(* IEC 61131-3 sources: rusty/tests/lit/single/polymorphism/fnptr, 14 files *)

(* ---- function_block_call_explicit_arguments.st ---- *)
// RUN: %COMPILE %s && %RUN | %CHECK %s

TYPE Position2D:
    STRUCT
        x: DINT;
        y: DINT;
    END_STRUCT
END_TYPE

FUNCTION_BLOCK FbA
    VAR
        localState: DINT := 0;
    END_VAR

    VAR_INPUT
        in1: DINT;
        in2: STRING;
        in3: Position2D;
        in4: ARRAY[1..2] OF STRING;
        in5: ARRAY[1..2] OF Position2D;
    END_VAR

    VAR_OUTPUT
        out1: DINT;
        out2: STRING;
        out3: Position2D;
        out4: ARRAY[1..2] OF STRING;
        out5: ARRAY[1..2] OF Position2D;
    END_VAR

    VAR_IN_OUT
        inout1: DINT;
        inout2: STRING;
        inout3: Position2D;
        inout4: ARRAY[1..2] OF STRING;
        inout5: ARRAY[1..2] OF Position2D;
    END_VAR

    METHOD increaseLocalState
        localState := localState + 1;
    END_METHOD

    printf('localState = %d$N', localState);

    printf('in1 = %d$N', in1);
    printf('in2 = %s$N', ADR(in2));
    printf('in3 = (%d, %d)$N', in3.x, in3.y);
    printf('in4 = [%s, %s]$N', ADR(in4[1]), ADR(in4[2]));
    printf('in5 = [(%d, %d), (%d, %d)]$N', in5[1].x, in5[1].y, in5[2].x, in5[2].y);

    printf('inout1 = %d$N', inout1);
    printf('inout2 = %s$N', ADR(inout2));
    printf('inout3 = (%d, %d)$N', inout3.x, inout3.y);
    printf('inout4 = [%s, %s]$N', ADR(inout4[1]), ADR(inout4[2]));
    printf('inout5 = [(%d, %d), (%d, %d)]$N', inout5[1].x, inout5[1].y, inout5[2].x, inout5[2].y);

    out1 := 55;
    out2 := 'sixty';
    out3.x := 65;
    out3.y := 70;
    out4[1] := 'seventy-five';
    out4[2] := 'eighty';
    out5[1].x := 85;
    out5[1].y := 90;
    out5[2].x := 95;
    out5[2].y := 100;

    inout1 := 105;
    inout2 := 'one-hundred-ten';
    inout3.x := 115;
    inout3.y := 120;
    inout4[1] := 'one-hundred-twenty-five';
    inout4[2] := 'one-hundred-thirty';
    inout5[1].x := 135;
    inout5[1].y := 140;
    inout5[2].x := 145;
    inout5[2].y := 150;
END_FUNCTION_BLOCK

FUNCTION main
    VAR
        instanceFbA: FbA;
        bodyPtr: __FPOINTER FbA := ADR(FbA);

        localIn1: DINT;
        localIn2: STRING;
        localIn3: Position2D;
        localIn4: ARRAY[1..2] OF STRING;
        localIn5: ARRAY[1..2] OF Position2D;

        localOut1: DINT;
        localOut2: STRING;
        localOut3: Position2D;
        localOut4: ARRAY[1..2] OF STRING;
        localOut5: ARRAY[1..2] OF Position2D;

        localInout1: DINT;
        localInout2: STRING;
        localInout3: Position2D;
        localInout4: ARRAY[1..2] OF STRING;
        localInout5: ARRAY[1..2] OF Position2D;
    END_VAR

    localIn3.x := 15;
    localIn3.y := 20;
    localIn4[1] := 'twenty-five';
    localIn4[2] := 'thirty';
    localIn5[1].x := 35;
    localIn5[1].y := 40;
    localIn5[2].x := 45;
    localIn5[2].y := 50;

    instanceFbA.increaseLocalState();

    // Partially initialized
    // localState = 1
    // CHECK: in1 = 0
    // CHECK: in2 =
    // CHECK: in3 = (15, 20)
    // CHECK: in4 = [twenty-five, thirty]
    // CHECK: in5 = [(35, 40), (45, 50)]
    // CHECK: inout1 = 0
    // CHECK: inout2 =
    // CHECK: inout3 = (0, 0)
    // CHECK: inout4 = [, ]
    // CHECK: inout5 = [(0, 0), (0, 0)]
    bodyPtr^(
        instanceFbA,
        inout5 := localInout5,
        in1 := localIn1,
        in2 := localIn2,
        in3 := localIn3,
        in4 := localIn4,
        in5 := localIn5,
        out1 => localOut1,
        out2 => localOut2,
        out3 => localOut3,
        out4 => localOut4,
        out5 => localOut5,
        inout1 := localInout1,
        inout2 := localInout2,
        inout3 := localInout3,
        inout4 := localInout4
    );

    // Locally, these should not be modified even if touched by the function block because they are passed by value
    // CHECK: localIn1 = 0
    // CHECK: localIn2 =
    // CHECK: localIn3 = (15, 20)
    // CHECK: localIn4 = [twenty-five, thirty]
    // CHECK: localIn5 = [(35, 40), (45, 50)]
    printf('localIn1 = %d$N', localIn1);
    printf('localIn2 = %s$N', ADR(localIn2));
    printf('localIn3 = (%d, %d)$N', localIn3.x, localIn3.y);
    printf('localIn4 = [%s, %s]$N', ADR(localIn4[1]), ADR(localIn4[2]));
    printf('localIn5 = [(%d, %d), (%d, %d)]$N', localIn5[1].x, localIn5[1].y, localIn5[2].x, localIn5[2].y);

    // Locally, these should be modified because they are passed by reference (not really but kind of)
    // CHECK: localOut1 = 55
    // CHECK: localOut2 = sixty
    // CHECK: localOut3 = (65, 70)
    // CHECK: localOut4 = [seventy-five, eighty]
    // CHECK: localOut5 = [(85, 90), (95, 100)]
    printf('localOut1 = %d$N', localOut1);
    printf('localOut2 = %s$N', ADR(localOut2));
    printf('localOut3 = (%d, %d)$N', localOut3.x, localOut3.y);
    printf('localOut4 = [%s, %s]$N', ADR(localOut4[1]), ADR(localOut4[2]));
    printf('localOut5 = [(%d, %d), (%d, %d)]$N', localOut5[1].x, localOut5[1].y, localOut5[2].x, localOut5[2].y);

    // Locally, these should be modified because they are passed by reference
    // CHECK: localInout1 = 105
    // CHECK: localInout2 = one-hundred-ten
    // CHECK: localInout3 = (115, 120)
    // CHECK: localInout4 = [one-hundred-twenty-five, one-hundred-thirty]
    // CHECK: localInout5 = [(135, 140), (145, 150)]
    printf('localInout1 = %d$N', localInout1);
    printf('localInout2 = %s$N', ADR(localInout2));
    printf('localInout3 = (%d, %d)$N', localInout3.x, localInout3.y);
    printf('localInout4 = [%s, %s]$N', ADR(localInout4[1]), ADR(localInout4[2]));
    printf('localInout5 = [(%d, %d), (%d, %d)]$N', localInout5[1].x, localInout5[1].y, localInout5[2].x, localInout5[2].y);
END_FUNCTION

(* ---- function_block_call_implicit_arguments.st ---- *)
// RUN: %COMPILE %s && %RUN | %CHECK %s

TYPE Position2D:
    STRUCT
        x: DINT;
        y: DINT;
    END_STRUCT
END_TYPE

FUNCTION_BLOCK FbA
    VAR
        localState: DINT := 0;
    END_VAR

    VAR_INPUT
        in1: DINT;
        in2: STRING;
        in3: Position2D;
        in4: ARRAY[1..2] OF STRING;
        in5: ARRAY[1..2] OF Position2D;
    END_VAR

    VAR_OUTPUT
        out1: DINT;
        out2: STRING;
        out3: Position2D;
        out4: ARRAY[1..2] OF STRING;
        out5: ARRAY[1..2] OF Position2D;
    END_VAR

    VAR_IN_OUT
        inout1: DINT;
        inout2: STRING;
        inout3: Position2D;
        inout4: ARRAY[1..2] OF STRING;
        inout5: ARRAY[1..2] OF Position2D;
    END_VAR

    METHOD increaseLocalState
        localState := localState + 1;
    END_METHOD

    printf('localState = %d$N', localState);

    printf('in1 = %d$N', in1);
    printf('in2 = %s$N', ADR(in2));
    printf('in3 = (%d, %d)$N', in3.x, in3.y);
    printf('in4 = [%s, %s]$N', ADR(in4[1]), ADR(in4[2]));
    printf('in5 = [(%d, %d), (%d, %d)]$N', in5[1].x, in5[1].y, in5[2].x, in5[2].y);

    printf('inout1 = %d$N', inout1);
    printf('inout2 = %s$N', ADR(inout2));
    printf('inout3 = (%d, %d)$N', inout3.x, inout3.y);
    printf('inout4 = [%s, %s]$N', ADR(inout4[1]), ADR(inout4[2]));
    printf('inout5 = [(%d, %d), (%d, %d)]$N', inout5[1].x, inout5[1].y, inout5[2].x, inout5[2].y);

    out1 := 55;
    out2 := 'sixty';
    out3.x := 65;
    out3.y := 70;
    out4[1] := 'seventy-five';
    out4[2] := 'eighty';
    out5[1].x := 85;
    out5[1].y := 90;
    out5[2].x := 95;
    out5[2].y := 100;

    inout1 := 105;
    inout2 := 'one-hundred-ten';
    inout3.x := 115;
    inout3.y := 120;
    inout4[1] := 'one-hundred-twenty-five';
    inout4[2] := 'one-hundred-thirty';
    inout5[1].x := 135;
    inout5[1].y := 140;
    inout5[2].x := 145;
    inout5[2].y := 150;
END_FUNCTION_BLOCK

FUNCTION main
    VAR
        instanceFbA: FbA;
        bodyPtr: __FPOINTER FbA := ADR(FbA);

        localIn1: DINT;
        localIn2: STRING;
        localIn3: Position2D;
        localIn4: ARRAY[1..2] OF STRING;
        localIn5: ARRAY[1..2] OF Position2D;

        localOut1: DINT;
        localOut2: STRING;
        localOut3: Position2D;
        localOut4: ARRAY[1..2] OF STRING;
        localOut5: ARRAY[1..2] OF Position2D;

        localInout1: DINT;
        localInout2: STRING;
        localInout3: Position2D;
        localInout4: ARRAY[1..2] OF STRING;
        localInout5: ARRAY[1..2] OF Position2D;
    END_VAR

    localIn3.x := 15;
    localIn3.y := 20;
    localIn4[1] := 'twenty-five';
    localIn4[2] := 'thirty';
    localIn5[1].x := 35;
    localIn5[1].y := 40;
    localIn5[2].x := 45;
    localIn5[2].y := 50;

    instanceFbA.increaseLocalState();

    // Partially initialized
    // localState = 1
    // CHECK: in1 = 0
    // CHECK: in2 =
    // CHECK: in3 = (15, 20)
    // CHECK: in4 = [twenty-five, thirty]
    // CHECK: in5 = [(35, 40), (45, 50)]
    // CHECK: inout1 = 0
    // CHECK: inout2 =
    // CHECK: inout3 = (0, 0)
    // CHECK: inout4 = [, ]
    // CHECK: inout5 = [(0, 0), (0, 0)]
    bodyPtr^(
        instanceFbA,
        localIn1,
        localIn2,
        localIn3,
        localIn4,
        localIn5,
        localOut1,
        localOut2,
        localOut3,
        localOut4,
        localOut5,
        localInout1,
        localInout2,
        localInout3,
        localInout4,
        localInout5
    );

    // Locally, these should not be modified even if touched by the function block because they are passed by value
    // CHECK: localIn1 = 0
    // CHECK: localIn2 =
    // CHECK: localIn3 = (15, 20)
    // CHECK: localIn4 = [twenty-five, thirty]
    // CHECK: localIn5 = [(35, 40), (45, 50)]
    printf('localIn1 = %d$N', localIn1);
    printf('localIn2 = %s$N', ADR(localIn2));
    printf('localIn3 = (%d, %d)$N', localIn3.x, localIn3.y);
    printf('localIn4 = [%s, %s]$N', ADR(localIn4[1]), ADR(localIn4[2]));
    printf('localIn5 = [(%d, %d), (%d, %d)]$N', localIn5[1].x, localIn5[1].y, localIn5[2].x, localIn5[2].y);

    // Locally, these should be modified because they are passed by reference (not really but kind of)
    // CHECK: localOut1 = 55
    // CHECK: localOut2 = sixty
    // CHECK: localOut3 = (65, 70)
    // CHECK: localOut4 = [seventy-five, eighty]
    // CHECK: localOut5 = [(85, 90), (95, 100)]
    printf('localOut1 = %d$N', localOut1);
    printf('localOut2 = %s$N', ADR(localOut2));
    printf('localOut3 = (%d, %d)$N', localOut3.x, localOut3.y);
    printf('localOut4 = [%s, %s]$N', ADR(localOut4[1]), ADR(localOut4[2]));
    printf('localOut5 = [(%d, %d), (%d, %d)]$N', localOut5[1].x, localOut5[1].y, localOut5[2].x, localOut5[2].y);

    // Locally, these should be modified because they are passed by reference
    // CHECK: localInout1 = 105
    // CHECK: localInout2 = one-hundred-ten
    // CHECK: localInout3 = (115, 120)
    // CHECK: localInout4 = [one-hundred-twenty-five, one-hundred-thirty]
    // CHECK: localInout5 = [(135, 140), (145, 150)]
    printf('localInout1 = %d$N', localInout1);
    printf('localInout2 = %s$N', ADR(localInout2));
    printf('localInout3 = (%d, %d)$N', localInout3.x, localInout3.y);
    printf('localInout4 = [%s, %s]$N', ADR(localInout4[1]), ADR(localInout4[2]));
    printf('localInout5 = [(%d, %d), (%d, %d)]$N', localInout5[1].x, localInout5[1].y, localInout5[2].x, localInout5[2].y);
END_FUNCTION

(* ---- function_block_call_local_variables.st ---- *)
// RUN: %COMPILE %s && %RUN | %CHECK %s

TYPE Position: STRUCT
        x: DINT;
        y: DINT;
    END_STRUCT
END_TYPE

FUNCTION_BLOCK A
    VAR
        localStateInt: DINT;
        localStateString: STRING;
        localStatePosition: Position;
        localStateStringArray: ARRAY[1..2] OF STRING;
        localStatePositionArray: ARRAY[1..2] OF Position;
    END_VAR

    METHOD printState
        printf('A::printState: localStateInt = %d$N', localStateInt);
        printf('A::printState: localStateString = %s$N', ADR(localStateString));
        printf('A::printState: localStatePosition = (%d, %d)$N', localStatePosition.x, localStatePosition.y);
        printf('A::printState: localStateStringArray[1] = %s$N', ADR(localStateStringArray[1]));
        printf('A::printState: localStateStringArray[2] = %s$N', ADR(localStateStringArray[2]));
        printf('A::printState: localStatePositionArray[1] = (%d, %d)$N', localStatePositionArray[1].x, localStatePositionArray[1].y);
        printf('A::printState: localStatePositionArray[2] = (%d, %d)$N', localStatePositionArray[2].x, localStatePositionArray[2].y);
    END_METHOD

    METHOD reset
        THIS^();
    END_METHOD

    // Init
    localStateInt := 5;
    localStateString := 'ten';
    localStatePosition.x := 15;
    localStatePosition.y := 20;
    localStateStringArray[1] := 'twenty-five';
    localStateStringArray[2] := 'thirty';
    localStatePositionArray[1].x := 35;
    localStatePositionArray[1].y := 40;
    localStatePositionArray[2].x := 45;
    localStatePositionArray[2].y := 50;
END_FUNCTION_BLOCK

FUNCTION main
    VAR
        instanceA: A;
        fnPtrBody: __FPOINTER A := ADR(A);
    END_VAR

    // CHECK: A::printState: localStateInt = 0
    // CHECK: A::printState: localStateString =
    // CHECK: A::printState: localStatePosition = (0, 0)
    // CHECK: A::printState: localStateStringArray[1] =
    // CHECK: A::printState: localStateStringArray[2] =
    // CHECK: A::printState: localStatePositionArray[1] = (0, 0)
    // CHECK: A::printState: localStatePositionArray[2] = (0, 0)
    instanceA.printState();

    // CHECK: A::printState: localStateInt = 5
    // CHECK: A::printState: localStateString = ten
    // CHECK: A::printState: localStatePosition = (15, 20)
    // CHECK: A::printState: localStateStringArray[1] = twenty-five
    // CHECK: A::printState: localStateStringArray[2] = thirty
    // CHECK: A::printState: localStatePositionArray[1] = (35, 40)
    // CHECK: A::printState: localStatePositionArray[2] = (45, 50)
    fnPtrBody^(instanceA);
    instanceA.printState();
END_FUNCTION

(* ---- method_call.st ---- *)
// RUN: %COMPILE %s && %RUN | %CHECK %s

FUNCTION_BLOCK FbA
    VAR
        localState: DINT := 5;
    END_VAR

    METHOD increaseStateByOne
        localState := localState + 1;
        printf('FbA::increaseStateByOne: localState = %d$N', localState);
    END_METHOD

    METHOD increaseStateByArg
        VAR_INPUT
            in: DINT;
        END_VAR

        localState := localState + in;
        printf('FbA::increaseStateByArg: localState = %d$N', localState);
    END_METHOD
END_FUNCTION_BLOCK

FUNCTION main
    VAR
        instanceFbA: FbA;
        fnPtrIncreaseStateByOne: __FPOINTER FbA.increaseStateByOne := ADR(FbA.increaseStateByOne);
        fnPtrIncreaseStateByArg: __FPOINTER FbA.increaseStateByArg := ADR(FbA.increaseStateByArg);
    END_VAR

    // CHECK: FbA::increaseStateByOne: localState = 6
    // CHECK: FbA::increaseStateByArg: localState = 10
    fnPtrIncreaseStateByOne^(instanceFbA);
    fnPtrIncreaseStateByArg^(instanceFbA, 4);
END_FUNCTION

(* ---- method_call_aggregate_return.st ---- *)
// RUN: %COMPILE %s && %RUN | %CHECK %s

TYPE PositionWithExtraMetadata:
    STRUCT
        x: REAL;
        y: REAL;
        data: ARRAY[1..100] OF STRING;
    END_STRUCT
END_TYPE

FUNCTION_BLOCK FbA
    VAR
        localStruct: PositionWithExtraMetadata := (x := 1.0, y := 2.0, data := ['Data 1', 'Data 2', 'Data 3']);
        localStringArray: ARRAY[1..3] OF STRING := ['Value 1', 'Value 2', 'Value 3'];
        localStructArray: ARRAY[1..3] OF PositionWithExtraMetadata := [
            (x := 3.0, y := 4.0, data := ['Data 4', 'Data 5', 'Data 6']),
            (x := 5.0, y := 6.0, data := ['Data 7', 'Data 8', 'Data 9']),
            (x := 7.0, y := 8.0, data := ['Data 10', 'Data 11', 'Data 12'])
        ];
    END_VAR

    METHOD returnString: STRING
        returnString := 'FbA::returnString';
    END_METHOD

    METHOD returnStruct: PositionWithExtraMetadata
        returnStruct := localStruct;
    END_METHOD

    METHOD returnStringArray: ARRAY[1..3] OF STRING
        returnStringArray := localStringArray;
    END_METHOD

    METHOD returnStructArray: ARRAY[1..3] OF PositionWithExtraMetadata
        returnStructArray := localStructArray;
    END_METHOD
END_FUNCTION_BLOCK

FUNCTION main
    VAR
        instanceA: FbA;
        returnStringPtr: __FPOINTER FbA.returnString := ADR(instanceA.returnString);
        returnStructPtr: __FPOINTER FbA.returnStruct := ADR(instanceA.returnStruct);
        returnStringArrayPtr: __FPOINTER FbA.returnStringArray := ADR(instanceA.returnStringArray);
        returnStructArrayPtr: __FPOINTER FbA.returnStructArray := ADR(instanceA.returnStructArray);

        localReturnString: STRING;
        localReturnStruct: PositionWithExtraMetadata;
        localReturnStringArray: ARRAY[1..3] OF STRING;
        localReturnStructArray: ARRAY[1..3] OF PositionWithExtraMetadata;
    END_VAR

    // localReturnString := instanceA.returnString();
    // CHECK: localReturnString = FbA::returnString
    localReturnString := returnStringPtr^(instanceA);
    printf('localReturnString = %s$N', ADR(localReturnString));

    // localReturnStruct := instanceA.returnStruct();
    // CHECK: localReturnStruct.x = 1.000000
    // CHECK: localReturnStruct.y = 2.000000
    // CHECK: localReturnStruct.data[1] = Data 1
    // CHECK: localReturnStruct.data[2] = Data 2
    // CHECK: localReturnStruct.data[3] = Data 3
    localReturnStruct := returnStructPtr^(instanceA);
    printf('localReturnStruct.x = %f$N', localReturnStruct.x);
    printf('localReturnStruct.y = %f$N', localReturnStruct.y);
    printf('localReturnStruct.data[1] = %s$N', ADR(localReturnStruct.data[1]));
    printf('localReturnStruct.data[2] = %s$N', ADR(localReturnStruct.data[2]));
    printf('localReturnStruct.data[3] = %s$N', ADR(localReturnStruct.data[3]));

    // localReturnStringArray := instanceA.returnStringArray();
    // CHECK: localReturnStringArray[1] = Value 1
    // CHECK: localReturnStringArray[2] = Value 2
    // CHECK: localReturnStringArray[3] = Value 3
    localReturnStringArray := returnStringArrayPtr^(instanceA);
    printf('localReturnStringArray[1] = %s$N', ADR(localReturnStringArray[1]));
    printf('localReturnStringArray[2] = %s$N', ADR(localReturnStringArray[2]));
    printf('localReturnStringArray[3] = %s$N', ADR(localReturnStringArray[3]));

    // localReturnStructArray := instanceA.returnStructArray();
    // CHECK: localReturnStructArray[1].x = 3.000000
    // CHECK: localReturnStructArray[1].y = 4.000000
    // CHECK: localReturnStructArray[1].data[1] = Data 4
    // CHECK: localReturnStructArray[1].data[2] = Data 5
    // CHECK: localReturnStructArray[1].data[3] = Data 6
    // CHECK: localReturnStructArray[2].x = 5.000000
    // CHECK: localReturnStructArray[2].y = 6.000000
    // CHECK: localReturnStructArray[2].data[1] = Data 7
    // CHECK: localReturnStructArray[2].data[2] = Data 8
    // CHECK: localReturnStructArray[2].data[3] = Data 9
    // CHECK: localReturnStructArray[3].x = 7.000000
    // CHECK: localReturnStructArray[3].y = 8.000000
    // CHECK: localReturnStructArray[3].data[1] = Data 10
    // CHECK: localReturnStructArray[3].data[2] = Data 11
    // CHECK: localReturnStructArray[3].data[3] = Data 12
    localReturnStructArray := returnStructArrayPtr^(instanceA);
    printf('localReturnStructArray[1].x = %f$N', localReturnStructArray[1].x);
    printf('localReturnStructArray[1].y = %f$N', localReturnStructArray[1].y);
    printf('localReturnStructArray[1].data[1] = %s$N', ADR(localReturnStructArray[1].data[1]));
    printf('localReturnStructArray[1].data[2] = %s$N', ADR(localReturnStructArray[1].data[2]));
    printf('localReturnStructArray[1].data[3] = %s$N', ADR(localReturnStructArray[1].data[3]));
    printf('localReturnStructArray[2].x = %f$N', localReturnStructArray[2].x);
    printf('localReturnStructArray[2].y = %f$N', localReturnStructArray[2].y);
    printf('localReturnStructArray[2].data[1] = %s$N', ADR(localReturnStructArray[2].data[1]));
    printf('localReturnStructArray[2].data[2] = %s$N', ADR(localReturnStructArray[2].data[2]));
    printf('localReturnStructArray[2].data[3] = %s$N', ADR(localReturnStructArray[2].data[3]));
    printf('localReturnStructArray[3].x = %f$N', localReturnStructArray[3].x);
    printf('localReturnStructArray[3].y = %f$N', localReturnStructArray[3].y);
    printf('localReturnStructArray[3].data[1] = %s$N', ADR(localReturnStructArray[3].data[1]));
    printf('localReturnStructArray[3].data[2] = %s$N', ADR(localReturnStructArray[3].data[2]));
    printf('localReturnStructArray[3].data[3] = %s$N', ADR(localReturnStructArray[3].data[3]));
END_FUNCTION

(* ---- method_call_aggregate_return_by_inout.st ---- *)
// RUN: %COMPILE %s && %RUN | %CHECK %s

TYPE PositionWithExtraMetadata:
    STRUCT
        x: REAL;
        y: REAL;
        data: ARRAY[1..100] OF STRING;
    END_STRUCT
END_TYPE

FUNCTION_BLOCK FbA
    METHOD foo
        VAR_OUTPUT
            outString: STRING;
            outStruct: PositionWithExtraMetadata;
            outStructArray: ARRAY[1..5] OF PositionWithExtraMetadata;
        END_VAR

        outString := 'FbA::foo result';
        outStruct.x := 1.0;
        outStruct.y := 2.0;
        outStruct.data[1] := 'Data 1';
        outStruct.data[2] := 'Data 2';
        outStruct.data[3] := 'Data 3';
        outStructArray[1].x := 3.0;
        outStructArray[1].y := 4.0;
        outStructArray[1].data[1] := 'Data 4';
        outStructArray[1].data[2] := 'Data 5';
        outStructArray[1].data[3] := 'Data 6';
    END_METHOD
END_FUNCTION_BLOCK

FUNCTION main
    VAR
        fooPtr: __FPOINTER FbA.foo := ADR(FbA.foo);
        instanceA: FbA;
        localOutString: STRING;
        localOutStruct: PositionWithExtraMetadata;
        localOutStructArray: ARRAY[1..5] OF PositionWithExtraMetadata;
    END_VAR

    // CHECK: localOutString = FbA::foo result
    // CHECK: localOutStruct.x = 1.000000
    // CHECK: localOutStruct.y = 2.000000
    // CHECK: localOutStruct.data[1] = Data 1
    // CHECK: localOutStruct.data[2] = Data 2
    // CHECK: localOutStruct.data[3] = Data 3
    // CHECK: localOutStructArray[1].x = 3.000000
    // CHECK: localOutStructArray[1].y = 4.000000
    // CHECK: localOutStructArray[1].data[1] = Data 4
    // CHECK: localOutStructArray[1].data[2] = Data 5
    // CHECK: localOutStructArray[1].data[3] = Data 6
    fooPtr^(instanceA, outStructArray => localOutStructArray, outString => localOutString, outStruct => localOutStruct );
    printf('localOutString = %s$N', ADR(localOutString));
    printf('localOutStruct.x = %f$N', localOutStruct.x);
    printf('localOutStruct.y = %f$N', localOutStruct.y);
    printf('localOutStruct.data[1] = %s$N', ADR(localOutStruct.data[1]));
    printf('localOutStruct.data[2] = %s$N', ADR(localOutStruct.data[2]));
    printf('localOutStruct.data[3] = %s$N', ADR(localOutStruct.data[3]));
    printf('localOutStructArray[1].x = %f$N', localOutStructArray[1].x);
    printf('localOutStructArray[1].y = %f$N', localOutStructArray[1].y);
    printf('localOutStructArray[1].data[1] = %s$N', ADR(localOutStructArray[1].data[1]));
    printf('localOutStructArray[1].data[2] = %s$N', ADR(localOutStructArray[1].data[2]));
    printf('localOutStructArray[1].data[3] = %s$N', ADR(localOutStructArray[1].data[3]));
END_FUNCTION

(* ---- method_call_aggregate_return_by_output.st ---- *)
// RUN: %COMPILE %s && %RUN | %CHECK %s

TYPE PositionWithExtraMetadata:
    STRUCT
        x: REAL;
        y: REAL;
        data: ARRAY[1..100] OF STRING;
    END_STRUCT
END_TYPE

FUNCTION_BLOCK FbA
    METHOD foo
        VAR_OUTPUT
            outString: STRING;
            outStruct: PositionWithExtraMetadata;
            outStringArray: ARRAY[1..5] OF STRING;
            outStructArray: ARRAY[1..5] OF PositionWithExtraMetadata;
        END_VAR

        outString := 'FbA::foo result';
        outStruct.x := 1.0;
        outStruct.y := 2.0;
        outStruct.data[1] := 'Data 1';
        outStruct.data[2] := 'Data 2';
        outStruct.data[3] := 'Data 3';
        outStringArray[1] := 'Data 4';
        outStringArray[2] := 'Data 5';
        outStringArray[3] := 'Data 6';
        outStructArray[1].x := 3.0;
        outStructArray[1].y := 4.0;
        outStructArray[1].data[1] := 'Data 7';
        outStructArray[1].data[2] := 'Data 8';
        outStructArray[1].data[3] := 'Data 9';
    END_METHOD
END_FUNCTION_BLOCK

FUNCTION main
    VAR
        fooPtr: __FPOINTER FbA.foo := ADR(FbA.foo);
        instanceA: FbA;
        localOutString: STRING;
        localOutStruct: PositionWithExtraMetadata;
        localOutStringArray: ARRAY[1..5] OF STRING;
        localOutStructArray: ARRAY[1..5] OF PositionWithExtraMetadata;
    END_VAR

    // CHECK: localOutString = FbA::foo result
    // CHECK: localOutStruct.x = 1.000000
    // CHECK: localOutStruct.y = 2.000000
    // CHECK: localOutStruct.data[1] = Data 1
    // CHECK: localOutStruct.data[2] = Data 2
    // CHECK: localOutStruct.data[3] = Data 3
    // CHECK: localOutStringArray[1] = Data 4
    // CHECK: localOutStringArray[2] = Data 5
    // CHECK: localOutStringArray[3] = Data 6
    // CHECK: localOutStructArray[1].x = 3.000000
    // CHECK: localOutStructArray[1].y = 4.000000
    // CHECK: localOutStructArray[1].data[1] = Data 7
    // CHECK: localOutStructArray[1].data[2] = Data 8
    // CHECK: localOutStructArray[1].data[3] = Data 9
    fooPtr^(instanceA, outStructArray => localOutStructArray, outString => localOutString, outStruct => localOutStruct, outStringArray => localOutStringArray);
    printf('localOutString = %s$N', ADR(localOutString));
    printf('localOutStruct.x = %f$N', localOutStruct.x);
    printf('localOutStruct.y = %f$N', localOutStruct.y);
    printf('localOutStruct.data[1] = %s$N', ADR(localOutStruct.data[1]));
    printf('localOutStruct.data[2] = %s$N', ADR(localOutStruct.data[2]));
    printf('localOutStruct.data[3] = %s$N', ADR(localOutStruct.data[3]));
    printf('localOutStringArray[1] = %s$N', ADR(localOutStringArray[1]));
    printf('localOutStringArray[2] = %s$N', ADR(localOutStringArray[2]));
    printf('localOutStringArray[3] = %s$N', ADR(localOutStringArray[3]));
    printf('localOutStructArray[1].x = %f$N', localOutStructArray[1].x);
    printf('localOutStructArray[1].y = %f$N', localOutStructArray[1].y);
    printf('localOutStructArray[1].data[1] = %s$N', ADR(localOutStructArray[1].data[1]));
    printf('localOutStructArray[1].data[2] = %s$N', ADR(localOutStructArray[1].data[2]));
    printf('localOutStructArray[1].data[3] = %s$N', ADR(localOutStructArray[1].data[3]));
END_FUNCTION

(* ---- method_call_by_void_pointer_cast.st ---- *)
// RUN: %COMPILE %s && %RUN | %CHECK %s

FUNCTION_BLOCK A
    METHOD printArgs
        VAR_INPUT
            message: STRING;
            value: DINT;
        END_VAR

        printf('%s %d$N', ADR(message), value);
    END_METHOD
END_FUNCTION_BLOCK

TYPE FnTable:
    STRUCT
        printArgs: __FPOINTER A.printArgs := ADR(A.printArgs);
    END_STRUCT
END_TYPE

VAR_GLOBAL
    fnTableInstance: FnTable;
END_VAR

FUNCTION main
    VAR
        instanceA: A;
        fnTableRef: POINTER TO __VOID := ADR(fnTableInstance);
    END_VAR

    // Not a direct cast of a void pointer function but rather its virtual table, basically how the virtual
    // table is also accessed in lowered code (though the access happens in the POU rather than a local
    // variable in the main function)
    // CHECK: value = 5
    // CHECK: value = 5
    FnTable#(fnTableRef^).printArgs^(instanceA, 'value =', 5);
    FnTable#(fnTableRef^).printArgs^(instanceA, message := 'value =', value := 5);
END_FUNCTION

(* ---- method_call_inout_arguments.st ---- *)
// RUN: %COMPILE %s && %RUN | %CHECK %s

FUNCTION_BLOCK A
    METHOD inoutArguments
        VAR_IN_OUT
            inout1: DINT;
            inout2: DINT;
        END_VAR

        inout1 := 100;
        inout2 := 200;
        printf('A::inoutArguments: inout1 = %d, inout2 = %d$N', inout1, inout2);
    END_METHOD
END_FUNCTION_BLOCK

FUNCTION main
    VAR
        instanceA: A;
        localInOut1: DINT;
        localInOut2: DINT;

        fnPtrInOutArguments: __FPOINTER A.inoutArguments := ADR(A.inoutArguments);
    END_VAR

    // Explicit
    // CHECK: A::inoutArguments: inout1 = 100, inout2 = 200
    // CHECK: A::inoutArguments: inout1 = 100, inout2 = 200
    fnPtrInOutArguments^(instanceA, localInOut1, localInOut2);
    fnPtrInOutArguments^(instanceA, inout1 := localInOut1, inout2 := localInOut2);
END_FUNCTION

(* ---- method_call_input_arguments.st ---- *)
// RUN: %COMPILE %s && %RUN | %CHECK %s

FUNCTION_BLOCK A
    METHOD inputArguments
        VAR_INPUT
            in1: DINT;
            in2: DINT;
        END_VAR

        printf('A::inputArguments: in1 = %d, in2 = %d$N', in1, in2);
    END_METHOD
END_FUNCTION_BLOCK

FUNCTION main
    VAR
        instanceA: A;
        localOut1: DINT;
        localOut2: DINT;

        fnPtrInputArguments: __FPOINTER A.inputArguments := ADR(A.inputArguments);
    END_VAR

    // Implicit
    // CHECK: A::inputArguments: in1 = 5, in2 = 10
    // CHECK: A::inputArguments: in1 = 5, in2 = 10
    fnPtrInputArguments^(instanceA, 5, 10);
    fnPtrInputArguments^(instanceA, in1 := 5, in2 := 10);
END_FUNCTION

(* ---- method_call_output_arguments.st ---- *)
// RUN: %COMPILE %s && %RUN | %CHECK %s

FUNCTION_BLOCK A
    METHOD outputArguments
        VAR_OUTPUT
            out1: DINT;
            out2: DINT;
        END_VAR

        out1 := 100;
        out2 := 200;
        printf('A::outputArguments: out1 = %d, out2 = %d$N', out1, out2);
    END_METHOD
END_FUNCTION_BLOCK

FUNCTION main
    VAR
        instanceA: A;
        localOut1: DINT;
        localOut2: DINT;

        fnPtrOutputArguments: __FPOINTER A.outputArguments := ADR(A.outputArguments);
    END_VAR

    // Explicit
    // CHECK: A::outputArguments: out1 = 100, out2 = 200
    // CHECK: A::outputArguments: out1 = 100, out2 = 200
    fnPtrOutputArguments^(instanceA, localOut1, localOut2);
    fnPtrOutputArguments^(instanceA, out1 => localOut1, out2 => localOut2);
END_FUNCTION

(* ---- method_call_overridden.st ---- *)
// RUN: %COMPILE %s && %RUN | %CHECK %s

FUNCTION_BLOCK A
    VAR
        nameA: STRING := 'FUNCTION_BLOCK A';
    END_VAR

    METHOD printName
        printf('name = %s$N', ADR(nameA));
    END_METHOD
END_FUNCTION_BLOCK

FUNCTION_BLOCK B EXTENDS A
    VAR
        nameB: STRING := 'FUNCTION_BLOCK B';
    END_VAR

    METHOD printName
        printf('name = %s$N', ADR(nameB));
    END_METHOD
END_FUNCTION_BLOCK

FUNCTION_BLOCK C
    VAR
        nameC: STRING := 'FUNCTION_BLOCK C';
    END_VAR

    METHOD printName
        printf('name = %s$N', ADR(nameC));
    END_METHOD
END_FUNCTION_BLOCK

FUNCTION main
    VAR
        instanceA: A;
        instanceB: B;
        instanceC: C;
        fnPtrPrintName: __FPOINTER A.printName := ADR(A.printName);
    END_VAR

    // Ensure that child POUs can be passed to function pointers of both its own and parent POUs. When doing
    // so we expect a bitcast on these passed arguments to the (in this case) parent POU.
    // CHECK: name = FUNCTION_BLOCK A
    // CHECK: name = FUNCTION_BLOCK A
    fnPtrPrintName^(instanceA);
    fnPtrPrintName^(instanceB); // <- fnPtrPrintName points to A.printName but we pass instanceB which should be fine and result in a bitcast

    // To showcase, we could pass an UNRELATED instance to the function pointer. Because it expects something
    // along `void (%A)` in LLVM IR (no return type, no parameters) passing `instanceC` should result in a
    // bitcast to `A`. The function (printName) should then GEP the first member field because `name` is
    // positioned there, resulting in access onto `nameC` rather than `nameA` and therefore a complete
    // different result when compared with a child instance. Illustrated (without size information)
    // `type A = { string }` -- expanded --> `type A = { nameA }`
    // `type B = { A, string }` -- expanded --> `type B = { { nameA }, nameB }`
    // `type C = { string} -- expanded --> `type C = { nameC }`
    // That should explain why we get `FUNCTION_BLOCK A` when passing `instanceB` and also why we get
    // `FUNCTION_BLOCK C` when passing `instanceC`
    // CHECK: name = FUNCTION_BLOCK C
    fnPtrPrintName^(instanceC);
END_FUNCTION

(* ---- method_call_using_this.st ---- *)
// RUN: %COMPILE %s && %RUN | %CHECK %s

VAR_GLOBAL
    instanceVirtuaTableA: VirtualTableA;
    instanceVirtuaTableB: VirtualTableB;
    instanceVirtuaTableC: VirtualTableC;
END_VAR

TYPE VirtualTableA:
    STRUCT
        getName: __FPOINTER A.getName := ADR(A.getName);
        printName: __FPOINTER A.printName := ADR(A.printName);
    END_STRUCT
END_TYPE

TYPE VirtualTableB:
    STRUCT
        getName: __FPOINTER A.getName := ADR(A.getName);
        printName: __FPOINTER A.printName := ADR(A.printName);
    END_STRUCT
END_TYPE

TYPE VirtualTableC:
    STRUCT
        getName: __FPOINTER C.getName := ADR(C.getName);
        printName: __FPOINTER A.printName := ADR(A.printName);
    END_STRUCT
END_TYPE

FUNCTION_BLOCK A
    VAR
        vt: POINTER TO __VOID;
    END_VAR

    METHOD getName: STRING
        getName := 'A';
    END_METHOD

    METHOD printName
        VAR
            result: STRING;
        END_VAR

        printf('name = %s$N', ADR(VirtualTableA#(vt^).getName^(THIS^)));
    END_METHOD
END_FUNCTION_BLOCK

// Inherits A as is
FUNCTION_BLOCK B EXTENDS A
END_FUNCTION_BLOCK

// Overrides the `getName` method
FUNCTION_BLOCK C EXTENDS A
    METHOD getName: STRING
        getName := 'C';
    END_METHOD
END_FUNCTION_BLOCK

FUNCTION main
    VAR
        instanceA: A;
        instanceB: B;
        instanceC: C;
    END_VAR

    instanceA.vt := ADR(instanceVirtuaTableA);
    instanceB.vt := ADR(instanceVirtuaTableB);
    instanceC.vt := ADR(instanceVirtuaTableC);

    // The `printName` call will use the virtual table to call the correct `getName` method
    // CHECK: name = A
    // CHECK: name = A
    // CHECK: name = C
    instanceA.printName(); // base method, hence A
    instanceB.printName(); // B inherits A without overriding any methods, hence A
    instanceC.printName(); // C inherits A overriding the `getName` method, hence C
END_FUNCTION

(* ---- user_defined_polymorphism.st ---- *)
// RUN: %COMPILE %s && %RUN | %CHECK %s

// Virtual Table Definitions
TYPE UserVT_FbA:
    STRUCT
        printNumber: __FPOINTER FbA.printNumber := ADR(FbA.printNumber);
    END_STRUCT
END_TYPE

TYPE UserVT_FbB:
    STRUCT
        // No override, hence the ADR(FbA.<...>)
        printNumber: __FPOINTER FbA.printNumber := ADR(FbA.printNumber);
    END_STRUCT
END_TYPE

TYPE UserVT_FbC:
    STRUCT
        // override, hence the ADR(FbC.<...>)
        printNumber: __FPOINTER FbA.printNumber := ADR(FbC.printNumber);
    END_STRUCT
END_TYPE

// Virtual Table Instances
VAR_GLOBAL
    UserVT_FbA_instance: UserVT_FbA;
    UserVT_FbB_instance: UserVT_FbB;
    UserVT_FbC_instance: UserVT_FbC;
END_VAR

FUNCTION_BLOCK FbA
    VAR
        vt: POINTER TO __VOID;
        localStateA: DINT := 5;
    END_VAR

    METHOD printNumber
        VAR_INPUT
            in: DINT;
        END_VAR

        printf('FbA::printNumber: localStateA = %d, in = %d$N', localStateA, in);
    END_METHOD
END_FUNCTION_BLOCK

FUNCTION_BLOCK FbB EXTENDS FbA
    VAR
        localStateB: DINT := 10;
    END_VAR
END_FUNCTION_BLOCK

FUNCTION_BLOCK FbC EXTENDS FbA
    VAR
        localStateC: DINT := 15;
    END_VAR

    METHOD printNumber
        VAR_INPUT
            in: DINT;
        END_VAR

        printf('FbC::printNumber: localStateA = %d, localStateC = %d, in = %d$N', localStateA, localStateC, in);
    END_METHOD
END_FUNCTION_BLOCK

FUNCTION main
    VAR
        instanceFbA: FbA;
        instanceFbB: FbB;
        instanceFbC: FbC;
        refInstanceFbA: POINTER TO FbA;
    END_VAR

    // Virtual Table Initialization
    instanceFbA.vt := ADR(UserVT_FbA_instance);
    instanceFbB.vt := ADR(UserVT_FbB_instance);
    instanceFbC.vt := ADR(UserVT_FbC_instance);

    // CHECK: FbA::printNumber: localStateA = 5, in = 5
    refInstanceFbA := ADR(instanceFbA);
    UserVT_FbA#(refInstanceFbA^.vt^).printNumber^(refInstanceFbA^, 5);

    // CHECK: FbA::printNumber: localStateA = 5, in = 10
    refInstanceFbA := ADR(instanceFbB);
    UserVT_FbA#(refInstanceFbA^.vt^).printNumber^(refInstanceFbA^, 10);

    // CHECK: FbC::printNumber: localStateA = 5, localStateC = 15, in = 15
    refInstanceFbA := ADR(instanceFbC);
    UserVT_FbA#(refInstanceFbA^.vt^).printNumber^(refInstanceFbA^, 15);
END_FUNCTION
